// Generated by voz_llm_plc_agent
// Target: Siemens TIA Portal V18 - SCL external source
// Review and compile before any download to physical hardware.

FUNCTION_BLOCK "PLC_PRG"
{ S7_Optimized_Access := 'TRUE' }
VERSION : 0.1
VAR_INPUT
   I_Start : Bool := FALSE;
   I_Emergency : Bool := FALSE;
   I_Safety_Condition : Bool := FALSE;
END_VAR
VAR_OUTPUT
   Q_Alarm : Bool := FALSE;
   Q_Motor_Enable : Bool := FALSE;
END_VAR
VAR
   M_FaultLatch : Bool;
END_VAR
BEGIN
(* Arranque seguro con alarma si no existe la condicion habilitante *)
IF #I_Emergency THEN
    #Q_Motor_Enable := FALSE;
    #M_FaultLatch := TRUE;
ELSIF #I_Start AND NOT #I_Safety_Condition THEN
    #Q_Motor_Enable := FALSE;
    #M_FaultLatch := TRUE;
ELSIF #I_Start AND #I_Safety_Condition AND NOT #M_FaultLatch THEN
    #Q_Motor_Enable := TRUE;
END_IF;

IF FALSE AND NOT #I_Emergency THEN
    #M_FaultLatch := FALSE;
END_IF;

#Q_Alarm := #M_FaultLatch;
END_FUNCTION_BLOCK

DATA_BLOCK "DB_PLC_PRG"
{ S7_Optimized_Access := 'TRUE' }
VERSION : 0.1
NON_RETAIN
"PLC_PRG"
BEGIN
END_DATA_BLOCK

ORGANIZATION_BLOCK "Main"
{ S7_Optimized_Access := 'TRUE' }
VERSION : 0.1
BEGIN
   "DB_PLC_PRG"(
      I_Start := "I_Start",
      I_Emergency := "I_Emergency",
      I_Safety_Condition := "I_Safety_Condition",
      Q_Alarm => "Q_Alarm",
      Q_Motor_Enable => "Q_Motor_Enable"
   );
END_ORGANIZATION_BLOCK
